(* IEC 61131-3 sources: codesys-to-astra/src/POUs/F_C2aPad2, 2 files *)

(* ---- F_C2aPad2.decl.st ---- *)
// Назначение: число 0..99 -> две цифры с ведущим нулём (для форматов даты и времени FB_C2aRtc).
// Автор:      kr0nsch
// Версия:     0.1.0
// Документ:   docs/LIBMAP.md
FUNCTION F_C2aPad2 : STRING(2)
VAR_INPUT
    usiValue : USINT;   // значение 0..99
END_VAR

(* ---- F_C2aPad2.impl.st ---- *)
IF usiValue < 10 THEN  // lint:allow STL008 одна десятичная цифра
    F_C2aPad2 := CONCAT('0', USINT_TO_STRING(usiValue));
ELSE
    F_C2aPad2 := USINT_TO_STRING(usiValue MOD 100);  // lint:allow STL008 две десятичные цифры
END_IF
